Universal Robots URScript: T012_codellama_34b_baseline_rep2.urscript

def program():
    # Home the robot
    movej(p[0, 0, 0, 0, 0, 0], v=200.0)

    # Approach spot 1
    movel(p[0, 0, 0, 0, 0, 0], v=200.0)

    # Descend
